GLOBALCONSTANTS FastPacket (* Konstanten für Übungen 142/143 (NMEA 2000 Fast Packet) *)
  (* Standard: 61499-1; Description: Copyright (c) 2026 Meisterschulen am Ostbahnhof This program and the accompanying materials are made available under the terms of the Eclipse Public License 2.0 which is available at https://www.eclipse.org/legal/epl-2.0/ SPDX-License-Identifier: EPL-2.0 *)
  (* Version 1.0, 2026-11-17, Franz Höpfinger, Meisterschulen am Ostbahnhof, NMEA 2000 Fast Packet *)
  PACKAGE Uebungen::const::Uebung_140_149;
  VAR_GLOBAL CONSTANT
    PGN_FPT_PROP_00 : UDINT := UDINT#16#1FF00; (* 142/143: proprietäre Fast-Packet-PGN 0x1FF00 *)
  END_VAR
END_GLOBALCONSTANTS
